Fanuc KAREL source: kt00889.KL

-- PROVISIONAL review KL for V940-1; original PC SHA256 8963e2043ac9f6b553a0b81f7778d158dd22f203ff2bad0cf78a80116889e49d
-- Incomplete behavior may be omitted. Consult companion uncertainty JSON. Do not deploy.
PROGRAM KT00889
%NOLOCKGROUP
-- UNRESOLVED_DECL P1 type=000102
-- UNRESOLVED_DECL P2 type=000102
-- UNRESOLVED_DECL OUT type=000101
BEGIN
  -- V9_ZERO_TABLE_METADATA_HINT layout=0001; no indexed target words; source/name/runtime held
  -- UNRESOLVED_PC offsets 5-20; opcodes 2E,22,32,35
  -- UNRESOLVED_PC offsets 25-40; opcodes 2E,22,32,35
  -- UNRESOLVED_PC offsets 45-60; opcodes 2E,22,32,35
  -- UNRESOLVED_PC offsets 65-80; opcodes 2E,22,32,35
  -- UNRESOLVED_PC offsets 85-115; opcodes 27,27,49,7E,AD,76,7E,4A
  -- UNRESOLVED_PC offsets 120-124; opcodes 7F
END KT00889
